// TIA Portal V20 export
// export: Created 2026-10-12T16:46:22.8578297Z, ExportSetting WithDefaults, DisplayName Totally Integrated Automation Portal, DisplayVersion V20 Update 6, DisplayName TIA Portal Openness, DisplayVersion V20 Update 6, DisplayName TIA Portal Version Control Interface, DisplayVersion V20 Update 6, DisplayName SINAMICS Startdrive Advanced, DisplayVersion V20 SP1 Update 2, DisplayName SINAMICS Startdrive G110M, G120, G120C, G120D, G120P, G115D, DisplayVersion V20 SP1 Update 2, DisplayName SINAMICS Startdrive G130, G150, S120, S150, SINAMICS MV, G220, S200, S210, DisplayVersion V20 SP1 Update 2, DisplayName STEP 7 Professional, DisplayVersion V20 Update 6, DisplayName STEP 7 Safety, DisplayVersion V20 Update 2, DisplayName WinCC Basic/Comfort/Advanced, DisplayVersion V20 Update 6, DisplayName WinCC Professional, DisplayVersion V20 Update 6, DisplayName WinCC Unified, DisplayVersion V20 Update 6
TYPE "UDT_Bad_Rueckmeldung"
// stored: IsFailsafeCompliant false
   STRUCT
      WT { S7_SetPoint := 'True'} : Array[1..3] of "UDT_WT_Rueckmeldung";
      Ampel_Status : Int;
      Betriebsbereit : Bool;
      Heizung_1_Ist : Real;
      Heizung_1_Soll : Real;
      Heizung_2_Ist : Real;
      Heizung_2_Soll : Real;
      Pumpe_Laeuft : Bool;
      Pumpe_FU_Soll : Real;
      US_Laeuft : Bool;
      GR_Aktiv : Bool;
      GR_Strom_Ist : Real;
      GR_Spannung_Ist : Real;
      WB_X_Soll : Real;
      WB_Y_Soll : Real;
      Hand_Aktiv : Bool;
      Hand_Abgelehnt : Bool;
   END_STRUCT;
END_TYPE
